(* IEC 61131-3 sources: rusty/tests/lit/cfc/validation/unsupported_expression, 1 file *)

(* ---- functions.st ---- *)
FUNCTION f : DINT
    f := 1;
END_FUNCTION

FUNCTION isReady : BOOL
    isReady := TRUE;
END_FUNCTION
